SYSTEM FillerModule (* Module Filler, generated from its module specification *)
  (* Standard: 61499-2 *)
  APPLICATION Filler (* Module Filler on target pc (localhost, IO modbus; generated by modgen) *)
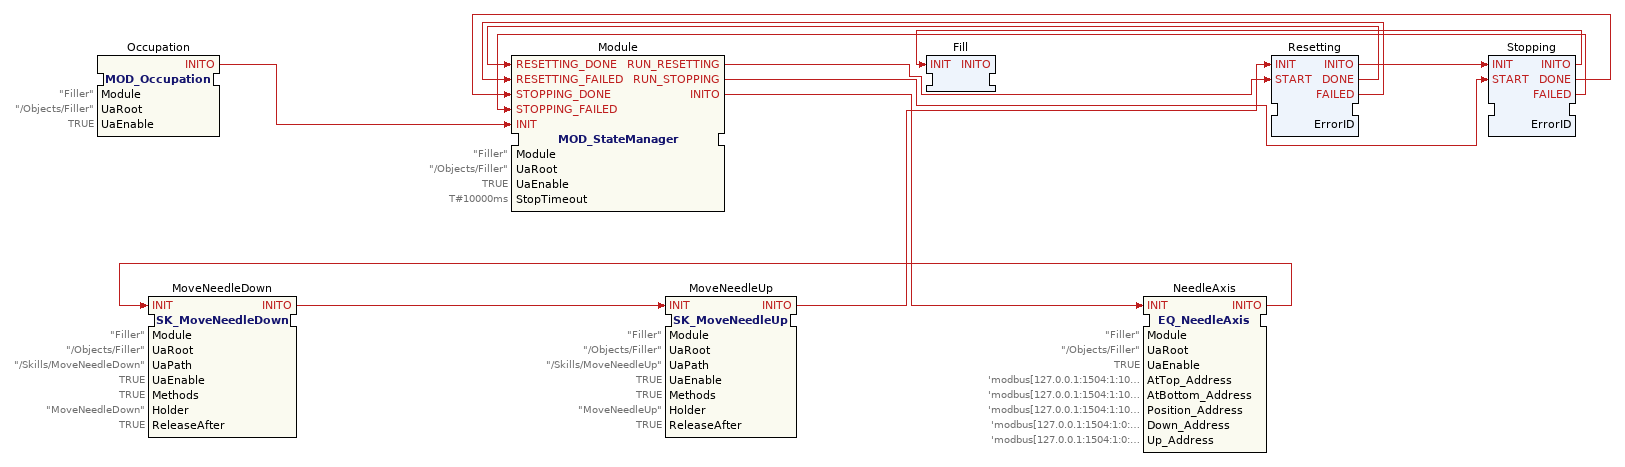
    (* Group ModuleLevel: Module level: occupation, PackML state manager, start-up and the target's IO lines *)
    (* Group ModuleLevelSkills: Module level skills: Control, Sequences (Execute, Stop) of skill primitives and Release; OPC UA /Skills/<name> *)
    (* Group Procedures: Procedures the module state manager runs while Resetting and Stopping *)
    (* Group SkillPrimitives: Skill primitives: one equipment command until a sensor or a time; OPC UA /Skills/<name> *)
    (* Group EquipmentIO: Equipment IO: the only owners of the IO points; skills send them output values over local channels *)
    FBS
      Occupation : modlib::MOD_Occupation(Module := "Filler", UaRoot := "/Objects/Filler", UaEnable := TRUE); (* Who may command the module. A client calls Occupy(Session) at /Objects/Filler/Occupation first; until it calls Release, only commands with that session id are accepted. Every block hears the owner on loc[Filler/owner]. *) {SET_ATTRIBUTE(GroupName, ModuleLevel)}
      Module : modlib::MOD_StateManager(Module := "Filler", UaRoot := "/Objects/Filler", UaEnable := TRUE, StopTimeout := T#10000ms); (* The module's PackML state. The owner calls Reset, Start, Stop, Abort or Clear at /Objects/Filler/Module; State is at /Objects/Filler/Module/State and on loc[Filler/state]. Reset runs the Resetting procedure, Stop the Stopping procedure; skills may be started only in Execute. *) {SET_ATTRIBUTE(GroupName, ModuleLevel)}
      NeedleAxis : filler::EQ_NeedleAxis(Module := "Filler", UaRoot := "/Objects/Filler", UaEnable := TRUE, AtTop_Address := 'modbus[127.0.0.1:1504:1:10:d0:]', AtBottom_Address := 'modbus[127.0.0.1:1504:1:10:d1:]', Position_Address := 'modbus[127.0.0.1:1504:1:10:i1:]', Down_Address := 'modbus[127.0.0.1:1504:1:0::c0]', Up_Address := 'modbus[127.0.0.1:1504:1:0::c2]'); (* Equipment NeedleAxis: Needle lift with down/up valves, end switches and a position sensor. The only block that touches its pins (AtTop = modbus[127.0.0.1:1504:1:10:d0:], AtBottom = modbus[127.0.0.1:1504:1:10:d1:], Position = modbus[127.0.0.1:1504:1:10:i1:], Down = modbus[127.0.0.1:1504:1:0::c0], Up = modbus[127.0.0.1:1504:1:0::c2]). Skills send it what to switch on loc[Filler/NeedleAxis/cmd]; it reports its inputs on loc[Filler/NeedleAxis/state] and at /Objects/Filler/Equipment/NeedleAxis. *) {SET_ATTRIBUTE(GroupName, EquipmentIO)}
      MoveNeedleDown : filler::SK_MoveNeedleDown(Module := "Filler", UaRoot := "/Objects/Filler", UaPath := "/Skills/MoveNeedleDown", UaEnable := TRUE, Methods := TRUE, Holder := "MoveNeedleDown", ReleaseAfter := TRUE); (* Skill MoveNeedleDown, offered on its own: Lower the needle to Distance mm below the top; the default is all the way down, using NeedleAxis. A client calls Start (with the parameters), Stop, Abort or Reset at /Objects/Filler/Skills/MoveNeedleDown; State, ErrorID, Parameters and Results are there too. *) {SET_ATTRIBUTE(GroupName, SkillPrimitives)}
      MoveNeedleUp : filler::SK_MoveNeedleUp(Module := "Filler", UaRoot := "/Objects/Filler", UaPath := "/Skills/MoveNeedleUp", UaEnable := TRUE, Methods := TRUE, Holder := "MoveNeedleUp", ReleaseAfter := TRUE); (* Skill MoveNeedleUp, offered on its own: Raise the needle to the top end switch, using NeedleAxis. A client calls Start (with the parameters), Stop, Abort or Reset at /Objects/Filler/Skills/MoveNeedleUp; State, ErrorID, Parameters and Results are there too. *) {SET_ATTRIBUTE(GroupName, SkillPrimitives)}
    END_FBS
    SUBAPPLICATION Resetting (* Procedure the module runs while Resetting *)
      {SET_ATTRIBUTE(GroupName, Procedures)}
      EVENT_INPUT
        INIT : EInit;
        START;
      END_EVENT
      EVENT_OUTPUT
        INITO : EInit;
        DONE;
        FAILED;
      END_EVENT
      VAR_OUTPUT
        ErrorID : UINT;
      END_VAR
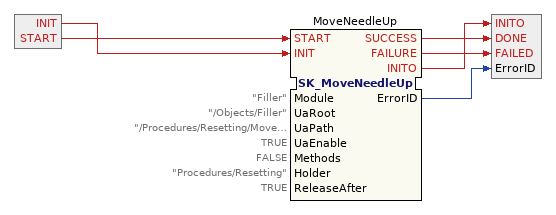
      FBS
        MoveNeedleUp : filler::SK_MoveNeedleUp(Module := "Filler", UaRoot := "/Objects/Filler", UaPath := "/Procedures/Resetting/MoveNeedleUp", UaEnable := TRUE, Methods := FALSE, Holder := "Procedures/Resetting", ReleaseAfter := TRUE); (* Step 1 of Resetting: runs the skill MoveNeedleUp. Its State and ErrorID are at /Objects/Filler/Procedures/Resetting/MoveNeedleUp; it keeps the equipment under the name Procedures/Resetting. *)
      END_FBS
      EVENT_CONNECTIONS
        START TO MoveNeedleUp.START;
        MoveNeedleUp.SUCCESS TO DONE;
        MoveNeedleUp.FAILURE TO FAILED;
        INIT TO MoveNeedleUp.INIT;
        MoveNeedleUp.INITO TO INITO;
      END_CONNECTIONS
      DATA_CONNECTIONS
        MoveNeedleUp.ErrorID TO ErrorID;
      END_CONNECTIONS
    END_SUBAPPLICATION
    SUBAPPLICATION Stopping (* Procedure the module runs while Stopping *)
      {SET_ATTRIBUTE(GroupName, Procedures)}
      EVENT_INPUT
        INIT : EInit;
        START;
      END_EVENT
      EVENT_OUTPUT
        INITO : EInit;
        DONE;
        FAILED;
      END_EVENT
      VAR_OUTPUT
        ErrorID : UINT;
      END_VAR
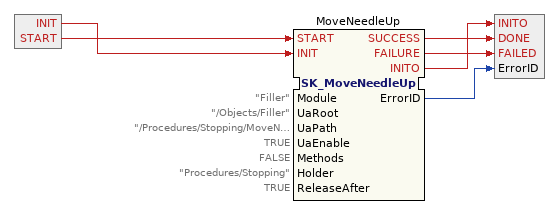
      FBS
        MoveNeedleUp : filler::SK_MoveNeedleUp(Module := "Filler", UaRoot := "/Objects/Filler", UaPath := "/Procedures/Stopping/MoveNeedleUp", UaEnable := TRUE, Methods := FALSE, Holder := "Procedures/Stopping", ReleaseAfter := TRUE); (* Step 1 of Stopping: runs the skill MoveNeedleUp. Its State and ErrorID are at /Objects/Filler/Procedures/Stopping/MoveNeedleUp; it keeps the equipment under the name Procedures/Stopping. *)
      END_FBS
      EVENT_CONNECTIONS
        START TO MoveNeedleUp.START;
        MoveNeedleUp.SUCCESS TO DONE;
        MoveNeedleUp.FAILURE TO FAILED;
        INIT TO MoveNeedleUp.INIT;
        MoveNeedleUp.INITO TO INITO;
      END_CONNECTIONS
      DATA_CONNECTIONS
        MoveNeedleUp.ErrorID TO ErrorID;
      END_CONNECTIONS
    END_SUBAPPLICATION
    SUBAPPLICATION Fill (* Module level skill Fill: Needle down to Depth and back up; a stop lifts the needle *)
      {SET_ATTRIBUTE(GroupName, ModuleLevelSkills)}
      EVENT_INPUT
        INIT : EInit;
      END_EVENT
      EVENT_OUTPUT
        INITO : EInit;
      END_EVENT
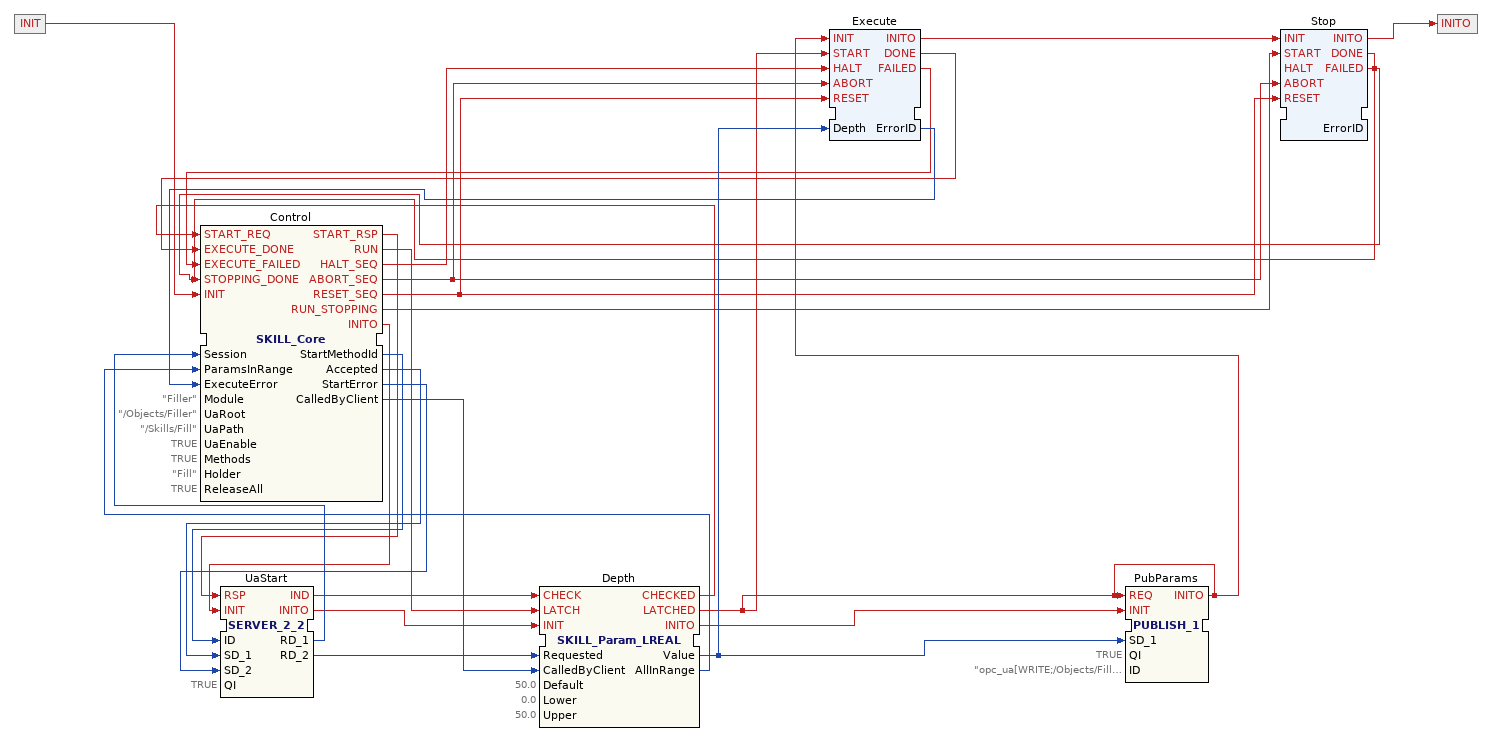
      (* Group Core: The skill's state machine: Stop, Abort, Reset, State and ErrorID over OPC UA; gives up everything the skill holds when a run ends *)
      (* Group Start: The Start method: one block per parameter (range check, value for this run), the values published *)
      (* Group Sequences: What the skill does: Execute, and Stop when it is interrupted; private skill primitives in order *)
      FBS
        Control : modlib::SKILL_Core(Module := "Filler", UaRoot := "/Objects/Filler", UaPath := "/Skills/Fill", UaEnable := TRUE, Methods := TRUE, Holder := "Fill", ReleaseAll := TRUE); (* The state machine of the skill Fill: checks a client's Start (occupation, module in Execute, not running, values in range), publishes State and ErrorID at /Objects/Filler/Skills/Fill, offers Stop, Abort and Reset there, starts Execute and runs Stop when the skill is stopped. *) {SET_ATTRIBUTE(GroupName, Core)}
        UaStart : iec61499::net::SERVER_2_2(QI := TRUE); (* The OPC UA method Start of Fill: a client's call (session id and parameters) arrives here; the parameters are checked, then Control answers Accepted or an error code. *) {SET_ATTRIBUTE(GroupName, Start)}
        Depth : modlib::SKILL_Param_LREAL(Default := 50.0, Lower := 0.0, Upper := 50.0); (* The parameter Depth of Fill: default 50.0 (Lower 0.0, Upper 50.0); checks a client's value, then holds it for the run and hands it to the steps. *) {SET_ATTRIBUTE(GroupName, Start)}
        PubParams : iec61499::net::PUBLISH_1(QI := TRUE, ID := "opc_ua[WRITE;/Objects/Filler/Skills/Fill/Parameters/Depth]"); (* Writes the parameters of the run to OPC UA: /Objects/Filler/Skills/Fill/Parameters/Depth *) {SET_ATTRIBUTE(GroupName, Start)}
      END_FBS
      SUBAPPLICATION Execute (* Fill: execute sequence *)
        {SET_ATTRIBUTE(GroupName, Sequences)}
        EVENT_INPUT
          INIT : EInit;
          START;
          HALT;
          ABORT;
          RESET;
        END_EVENT
        EVENT_OUTPUT
          INITO : EInit;
          DONE;
          FAILED;
        END_EVENT
        VAR_INPUT
          Depth : LREAL;
        END_VAR
        VAR_OUTPUT
          ErrorID : UINT;
        END_VAR
        FBS
          MoveNeedleDown : filler::SK_MoveNeedleDown(Module := "Filler", UaRoot := "/Objects/Filler", UaPath := "/Skills/Fill/Execute/MoveNeedleDown", UaEnable := TRUE, Methods := FALSE, Holder := "Fill", ReleaseAfter := FALSE); (* Step 1 of Fill / Execute: runs the skill MoveNeedleDown; Distance from Fill's Depth. Its State and ErrorID are at /Objects/Filler/Skills/Fill/Execute/MoveNeedleDown; it keeps the equipment under the name Fill. *)
          MoveNeedleUp : filler::SK_MoveNeedleUp(Module := "Filler", UaRoot := "/Objects/Filler", UaPath := "/Skills/Fill/Execute/MoveNeedleUp", UaEnable := TRUE, Methods := FALSE, Holder := "Fill", ReleaseAfter := FALSE); (* Step 2 of Fill / Execute: runs the skill MoveNeedleUp. Its State and ErrorID are at /Objects/Filler/Skills/Fill/Execute/MoveNeedleUp; it keeps the equipment under the name Fill. *)
          Fail1 : modlib::SKILL_FailMerge; (* Joins the failures of the steps into one (with its error code), so any step's failure ends the sequence. *)
        END_FBS
        EVENT_CONNECTIONS
          MoveNeedleDown.SUCCESS TO MoveNeedleUp.START;
          START TO MoveNeedleDown.START;
          MoveNeedleUp.SUCCESS TO DONE;
          MoveNeedleDown.FAILURE TO Fail1.FAIL_1;
          MoveNeedleUp.FAILURE TO Fail1.FAIL_2;
          Fail1.FAIL TO FAILED;
          INIT TO MoveNeedleDown.INIT;
          MoveNeedleUp.INITO TO INITO;
          MoveNeedleDown.INITO TO MoveNeedleUp.INIT;
          HALT TO MoveNeedleDown.HALT;
          HALT TO MoveNeedleUp.HALT;
          ABORT TO MoveNeedleDown.ABORT;
          ABORT TO MoveNeedleUp.ABORT;
          RESET TO MoveNeedleDown.RESET;
          RESET TO MoveNeedleUp.RESET;
        END_CONNECTIONS
        DATA_CONNECTIONS
          Depth TO MoveNeedleDown.Distance;
          MoveNeedleDown.ErrorID TO Fail1.Error1;
          MoveNeedleUp.ErrorID TO Fail1.Error2;
          Fail1.Error TO ErrorID;
        END_CONNECTIONS
      END_SUBAPPLICATION
      SUBAPPLICATION Stop (* Fill: stop sequence *)
        {SET_ATTRIBUTE(GroupName, Sequences)}
        EVENT_INPUT
          INIT : EInit;
          START;
          HALT;
          ABORT;
          RESET;
        END_EVENT
        EVENT_OUTPUT
          INITO : EInit;
          DONE;
          FAILED;
        END_EVENT
        VAR_OUTPUT
          ErrorID : UINT;
        END_VAR
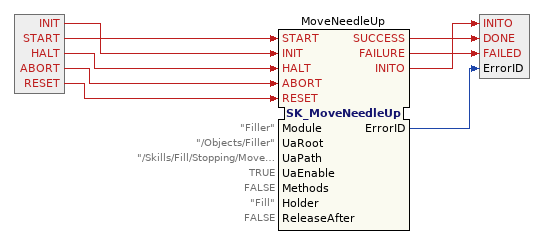
        FBS
          MoveNeedleUp : filler::SK_MoveNeedleUp(Module := "Filler", UaRoot := "/Objects/Filler", UaPath := "/Skills/Fill/Stopping/MoveNeedleUp", UaEnable := TRUE, Methods := FALSE, Holder := "Fill", ReleaseAfter := FALSE); (* Step 1 of Fill / Stop: runs the skill MoveNeedleUp. Its State and ErrorID are at /Objects/Filler/Skills/Fill/Stopping/MoveNeedleUp; it keeps the equipment under the name Fill. *)
        END_FBS
        EVENT_CONNECTIONS
          START TO MoveNeedleUp.START;
          MoveNeedleUp.SUCCESS TO DONE;
          MoveNeedleUp.FAILURE TO FAILED;
          INIT TO MoveNeedleUp.INIT;
          MoveNeedleUp.INITO TO INITO;
          HALT TO MoveNeedleUp.HALT;
          ABORT TO MoveNeedleUp.ABORT;
          RESET TO MoveNeedleUp.RESET;
        END_CONNECTIONS
        DATA_CONNECTIONS
          MoveNeedleUp.ErrorID TO ErrorID;
        END_CONNECTIONS
      END_SUBAPPLICATION
      EVENT_CONNECTIONS
        Control.START_RSP TO UaStart.RSP;
        UaStart.IND TO Depth.CHECK;
        Control.RUN TO Depth.LATCH;
        Depth.CHECKED TO Control.START_REQ;
        Depth.LATCHED TO PubParams.REQ;
        PubParams.INITO TO PubParams.REQ;
        Depth.LATCHED TO Execute.START;
        Control.HALT_SEQ TO Execute.HALT;
        Control.ABORT_SEQ TO Execute.ABORT;
        Control.RESET_SEQ TO Execute.RESET;
        Execute.DONE TO Control.EXECUTE_DONE;
        Execute.FAILED TO Control.EXECUTE_FAILED;
        Control.RUN_STOPPING TO Stop.START;
        Control.ABORT_SEQ TO Stop.ABORT;
        Control.RESET_SEQ TO Stop.RESET;
        Stop.DONE TO Control.STOPPING_DONE;
        Stop.FAILED TO Control.STOPPING_DONE;
        INIT TO Control.INIT;
        Control.INITO TO UaStart.INIT;
        UaStart.INITO TO Depth.INIT;
        Depth.INITO TO PubParams.INIT;
        PubParams.INITO TO Execute.INIT;
        Execute.INITO TO Stop.INIT;
        Stop.INITO TO INITO;
      END_CONNECTIONS
      DATA_CONNECTIONS
        Control.StartMethodId TO UaStart.ID;
        UaStart.RD_1 TO Control.Session;
        Control.Accepted TO UaStart.SD_1;
        Control.StartError TO UaStart.SD_2;
        UaStart.RD_2 TO Depth.Requested;
        Control.CalledByClient TO Depth.CalledByClient;
        Depth.Value TO PubParams.SD_1;
        Depth.AllInRange TO Control.ParamsInRange;
        Depth.Value TO Execute.Depth;
        Execute.ErrorID TO Control.ExecuteError;
      END_CONNECTIONS
    END_SUBAPPLICATION
    EVENT_CONNECTIONS
      Module.RUN_RESETTING TO Resetting.START;
      Resetting.DONE TO Module.RESETTING_DONE;
      Resetting.FAILED TO Module.RESETTING_FAILED;
      Module.RUN_STOPPING TO Stopping.START;
      Stopping.DONE TO Module.STOPPING_DONE;
      Stopping.FAILED TO Module.STOPPING_FAILED;
      Occupation.INITO TO Module.INIT;
      Module.INITO TO NeedleAxis.INIT;
      NeedleAxis.INITO TO MoveNeedleDown.INIT;
      MoveNeedleDown.INITO TO MoveNeedleUp.INIT;
      MoveNeedleUp.INITO TO Resetting.INIT;
      Resetting.INITO TO Stopping.INIT;
      Stopping.INITO TO Fill.INIT;
    END_CONNECTIONS
  END_APPLICATION
  APPLICATION Filler_pi (* Module Filler on target pi (filler-pi.invalid, IO gpio; generated by modgen) *)
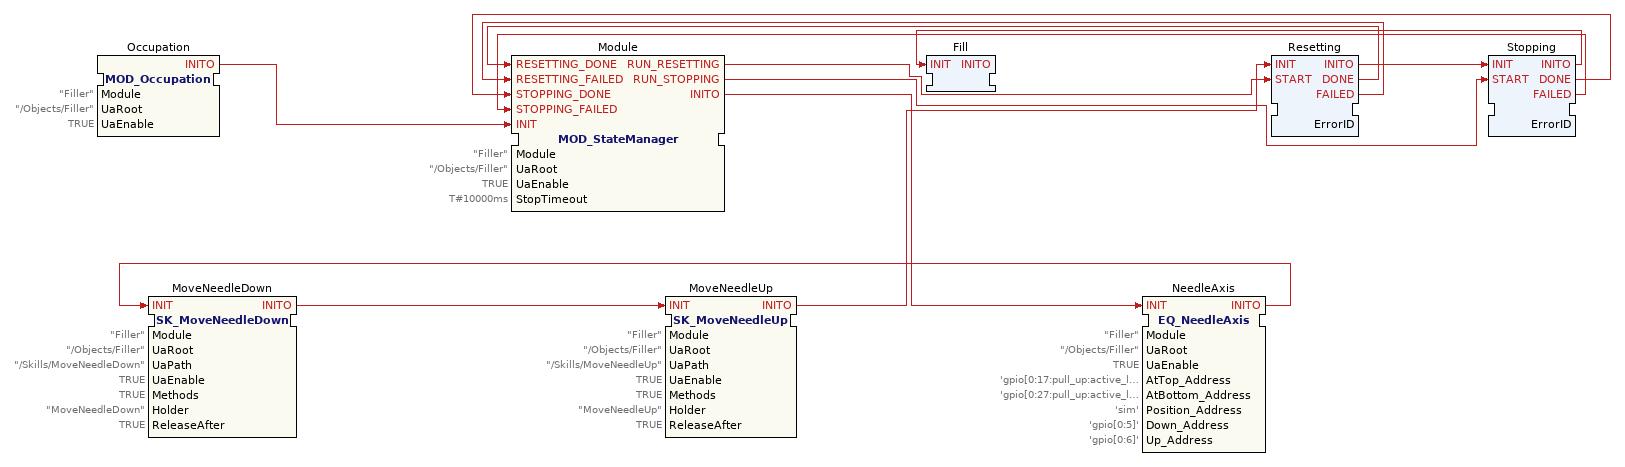
    (* Group ModuleLevel: Module level: occupation, PackML state manager, start-up and the target's IO lines *)
    (* Group ModuleLevelSkills: Module level skills: Control, Sequences (Execute, Stop) of skill primitives and Release; OPC UA /Skills/<name> *)
    (* Group Procedures: Procedures the module state manager runs while Resetting and Stopping *)
    (* Group SkillPrimitives: Skill primitives: one equipment command until a sensor or a time; OPC UA /Skills/<name> *)
    (* Group EquipmentIO: Equipment IO: the only owners of the IO points; skills send them output values over local channels *)
    FBS
      Occupation : modlib::MOD_Occupation(Module := "Filler", UaRoot := "/Objects/Filler", UaEnable := TRUE); (* Who may command the module. A client calls Occupy(Session) at /Objects/Filler/Occupation first; until it calls Release, only commands with that session id are accepted. Every block hears the owner on loc[Filler/owner]. *) {SET_ATTRIBUTE(GroupName, ModuleLevel)}
      Module : modlib::MOD_StateManager(Module := "Filler", UaRoot := "/Objects/Filler", UaEnable := TRUE, StopTimeout := T#10000ms); (* The module's PackML state. The owner calls Reset, Start, Stop, Abort or Clear at /Objects/Filler/Module; State is at /Objects/Filler/Module/State and on loc[Filler/state]. Reset runs the Resetting procedure, Stop the Stopping procedure; skills may be started only in Execute. *) {SET_ATTRIBUTE(GroupName, ModuleLevel)}
      NeedleAxis : filler::EQ_NeedleAxis(Module := "Filler", UaRoot := "/Objects/Filler", UaEnable := TRUE, AtTop_Address := 'gpio[0:17:pull_up:active_low]', AtBottom_Address := 'gpio[0:27:pull_up:active_low]', Position_Address := 'sim', Down_Address := 'gpio[0:5]', Up_Address := 'gpio[0:6]'); (* Equipment NeedleAxis: Needle lift with down/up valves, end switches and a position sensor. The only block that touches its pins (AtTop = gpio[0:17:pull_up:active_low], AtBottom = gpio[0:27:pull_up:active_low], Position = sim, Down = gpio[0:5], Up = gpio[0:6]). Skills send it what to switch on loc[Filler/NeedleAxis/cmd]; it reports its inputs on loc[Filler/NeedleAxis/state] and at /Objects/Filler/Equipment/NeedleAxis. *) {SET_ATTRIBUTE(GroupName, EquipmentIO)}
      MoveNeedleDown : filler::SK_MoveNeedleDown(Module := "Filler", UaRoot := "/Objects/Filler", UaPath := "/Skills/MoveNeedleDown", UaEnable := TRUE, Methods := TRUE, Holder := "MoveNeedleDown", ReleaseAfter := TRUE); (* Skill MoveNeedleDown, offered on its own: Lower the needle to Distance mm below the top; the default is all the way down, using NeedleAxis. A client calls Start (with the parameters), Stop, Abort or Reset at /Objects/Filler/Skills/MoveNeedleDown; State, ErrorID, Parameters and Results are there too. *) {SET_ATTRIBUTE(GroupName, SkillPrimitives)}
      MoveNeedleUp : filler::SK_MoveNeedleUp(Module := "Filler", UaRoot := "/Objects/Filler", UaPath := "/Skills/MoveNeedleUp", UaEnable := TRUE, Methods := TRUE, Holder := "MoveNeedleUp", ReleaseAfter := TRUE); (* Skill MoveNeedleUp, offered on its own: Raise the needle to the top end switch, using NeedleAxis. A client calls Start (with the parameters), Stop, Abort or Reset at /Objects/Filler/Skills/MoveNeedleUp; State, ErrorID, Parameters and Results are there too. *) {SET_ATTRIBUTE(GroupName, SkillPrimitives)}
    END_FBS
    SUBAPPLICATION Resetting (* Procedure the module runs while Resetting *)
      {SET_ATTRIBUTE(GroupName, Procedures)}
      EVENT_INPUT
        INIT : EInit;
        START;
      END_EVENT
      EVENT_OUTPUT
        INITO : EInit;
        DONE;
        FAILED;
      END_EVENT
      VAR_OUTPUT
        ErrorID : UINT;
      END_VAR
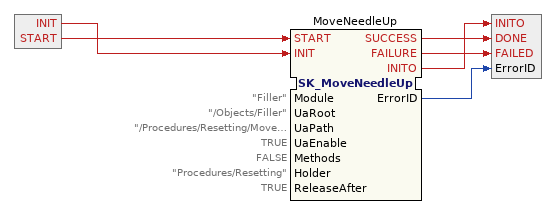
      FBS
        MoveNeedleUp : filler::SK_MoveNeedleUp(Module := "Filler", UaRoot := "/Objects/Filler", UaPath := "/Procedures/Resetting/MoveNeedleUp", UaEnable := TRUE, Methods := FALSE, Holder := "Procedures/Resetting", ReleaseAfter := TRUE); (* Step 1 of Resetting: runs the skill MoveNeedleUp. Its State and ErrorID are at /Objects/Filler/Procedures/Resetting/MoveNeedleUp; it keeps the equipment under the name Procedures/Resetting. *)
      END_FBS
      EVENT_CONNECTIONS
        START TO MoveNeedleUp.START;
        MoveNeedleUp.SUCCESS TO DONE;
        MoveNeedleUp.FAILURE TO FAILED;
        INIT TO MoveNeedleUp.INIT;
        MoveNeedleUp.INITO TO INITO;
      END_CONNECTIONS
      DATA_CONNECTIONS
        MoveNeedleUp.ErrorID TO ErrorID;
      END_CONNECTIONS
    END_SUBAPPLICATION
    SUBAPPLICATION Stopping (* Procedure the module runs while Stopping *)
      {SET_ATTRIBUTE(GroupName, Procedures)}
      EVENT_INPUT
        INIT : EInit;
        START;
      END_EVENT
      EVENT_OUTPUT
        INITO : EInit;
        DONE;
        FAILED;
      END_EVENT
      VAR_OUTPUT
        ErrorID : UINT;
      END_VAR
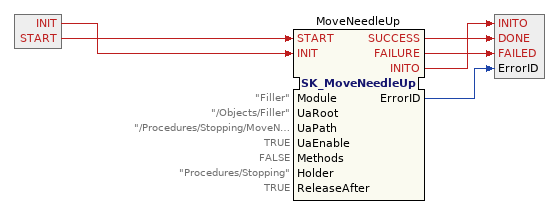
      FBS
        MoveNeedleUp : filler::SK_MoveNeedleUp(Module := "Filler", UaRoot := "/Objects/Filler", UaPath := "/Procedures/Stopping/MoveNeedleUp", UaEnable := TRUE, Methods := FALSE, Holder := "Procedures/Stopping", ReleaseAfter := TRUE); (* Step 1 of Stopping: runs the skill MoveNeedleUp. Its State and ErrorID are at /Objects/Filler/Procedures/Stopping/MoveNeedleUp; it keeps the equipment under the name Procedures/Stopping. *)
      END_FBS
      EVENT_CONNECTIONS
        START TO MoveNeedleUp.START;
        MoveNeedleUp.SUCCESS TO DONE;
        MoveNeedleUp.FAILURE TO FAILED;
        INIT TO MoveNeedleUp.INIT;
        MoveNeedleUp.INITO TO INITO;
      END_CONNECTIONS
      DATA_CONNECTIONS
        MoveNeedleUp.ErrorID TO ErrorID;
      END_CONNECTIONS
    END_SUBAPPLICATION
    SUBAPPLICATION Fill (* Module level skill Fill: Needle down to Depth and back up; a stop lifts the needle *)
      {SET_ATTRIBUTE(GroupName, ModuleLevelSkills)}
      EVENT_INPUT
        INIT : EInit;
      END_EVENT
      EVENT_OUTPUT
        INITO : EInit;
      END_EVENT
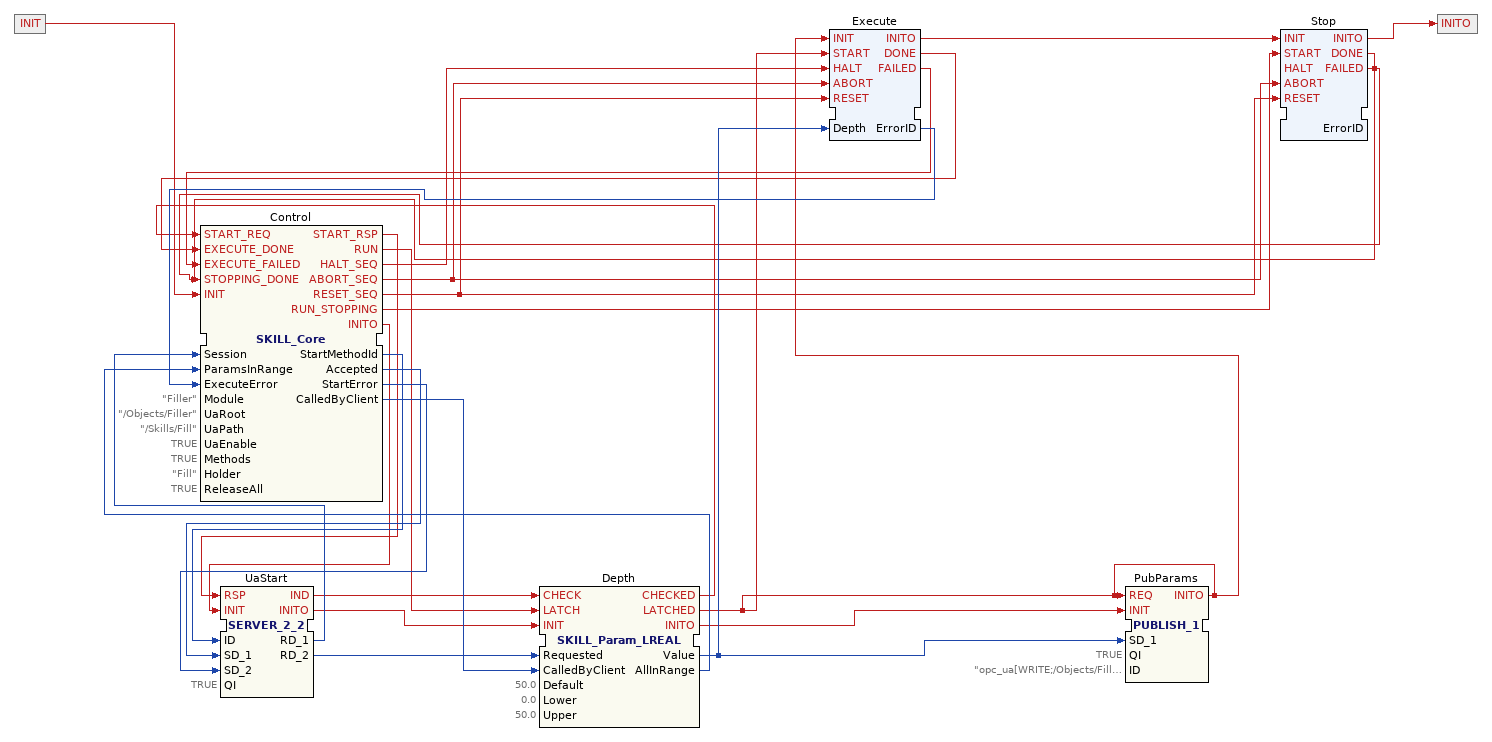
      (* Group Core: The skill's state machine: Stop, Abort, Reset, State and ErrorID over OPC UA; gives up everything the skill holds when a run ends *)
      (* Group Start: The Start method: one block per parameter (range check, value for this run), the values published *)
      (* Group Sequences: What the skill does: Execute, and Stop when it is interrupted; private skill primitives in order *)
      FBS
        Control : modlib::SKILL_Core(Module := "Filler", UaRoot := "/Objects/Filler", UaPath := "/Skills/Fill", UaEnable := TRUE, Methods := TRUE, Holder := "Fill", ReleaseAll := TRUE); (* The state machine of the skill Fill: checks a client's Start (occupation, module in Execute, not running, values in range), publishes State and ErrorID at /Objects/Filler/Skills/Fill, offers Stop, Abort and Reset there, starts Execute and runs Stop when the skill is stopped. *) {SET_ATTRIBUTE(GroupName, Core)}
        UaStart : iec61499::net::SERVER_2_2(QI := TRUE); (* The OPC UA method Start of Fill: a client's call (session id and parameters) arrives here; the parameters are checked, then Control answers Accepted or an error code. *) {SET_ATTRIBUTE(GroupName, Start)}
        Depth : modlib::SKILL_Param_LREAL(Default := 50.0, Lower := 0.0, Upper := 50.0); (* The parameter Depth of Fill: default 50.0 (Lower 0.0, Upper 50.0); checks a client's value, then holds it for the run and hands it to the steps. *) {SET_ATTRIBUTE(GroupName, Start)}
        PubParams : iec61499::net::PUBLISH_1(QI := TRUE, ID := "opc_ua[WRITE;/Objects/Filler/Skills/Fill/Parameters/Depth]"); (* Writes the parameters of the run to OPC UA: /Objects/Filler/Skills/Fill/Parameters/Depth *) {SET_ATTRIBUTE(GroupName, Start)}
      END_FBS
      SUBAPPLICATION Execute (* Fill: execute sequence *)
        {SET_ATTRIBUTE(GroupName, Sequences)}
        EVENT_INPUT
          INIT : EInit;
          START;
          HALT;
          ABORT;
          RESET;
        END_EVENT
        EVENT_OUTPUT
          INITO : EInit;
          DONE;
          FAILED;
        END_EVENT
        VAR_INPUT
          Depth : LREAL;
        END_VAR
        VAR_OUTPUT
          ErrorID : UINT;
        END_VAR
        FBS
          MoveNeedleDown : filler::SK_MoveNeedleDown(Module := "Filler", UaRoot := "/Objects/Filler", UaPath := "/Skills/Fill/Execute/MoveNeedleDown", UaEnable := TRUE, Methods := FALSE, Holder := "Fill", ReleaseAfter := FALSE); (* Step 1 of Fill / Execute: runs the skill MoveNeedleDown; Distance from Fill's Depth. Its State and ErrorID are at /Objects/Filler/Skills/Fill/Execute/MoveNeedleDown; it keeps the equipment under the name Fill. *)
          MoveNeedleUp : filler::SK_MoveNeedleUp(Module := "Filler", UaRoot := "/Objects/Filler", UaPath := "/Skills/Fill/Execute/MoveNeedleUp", UaEnable := TRUE, Methods := FALSE, Holder := "Fill", ReleaseAfter := FALSE); (* Step 2 of Fill / Execute: runs the skill MoveNeedleUp. Its State and ErrorID are at /Objects/Filler/Skills/Fill/Execute/MoveNeedleUp; it keeps the equipment under the name Fill. *)
          Fail1 : modlib::SKILL_FailMerge; (* Joins the failures of the steps into one (with its error code), so any step's failure ends the sequence. *)
        END_FBS
        EVENT_CONNECTIONS
          MoveNeedleDown.SUCCESS TO MoveNeedleUp.START;
          START TO MoveNeedleDown.START;
          MoveNeedleUp.SUCCESS TO DONE;
          MoveNeedleDown.FAILURE TO Fail1.FAIL_1;
          MoveNeedleUp.FAILURE TO Fail1.FAIL_2;
          Fail1.FAIL TO FAILED;
          INIT TO MoveNeedleDown.INIT;
          MoveNeedleUp.INITO TO INITO;
          MoveNeedleDown.INITO TO MoveNeedleUp.INIT;
          HALT TO MoveNeedleDown.HALT;
          HALT TO MoveNeedleUp.HALT;
          ABORT TO MoveNeedleDown.ABORT;
          ABORT TO MoveNeedleUp.ABORT;
          RESET TO MoveNeedleDown.RESET;
          RESET TO MoveNeedleUp.RESET;
        END_CONNECTIONS
        DATA_CONNECTIONS
          Depth TO MoveNeedleDown.Distance;
          MoveNeedleDown.ErrorID TO Fail1.Error1;
          MoveNeedleUp.ErrorID TO Fail1.Error2;
          Fail1.Error TO ErrorID;
        END_CONNECTIONS
      END_SUBAPPLICATION
      SUBAPPLICATION Stop (* Fill: stop sequence *)
        {SET_ATTRIBUTE(GroupName, Sequences)}
        EVENT_INPUT
          INIT : EInit;
          START;
          HALT;
          ABORT;
          RESET;
        END_EVENT
        EVENT_OUTPUT
          INITO : EInit;
          DONE;
          FAILED;
        END_EVENT
        VAR_OUTPUT
          ErrorID : UINT;
        END_VAR
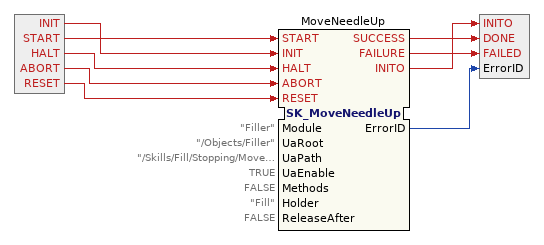
        FBS
          MoveNeedleUp : filler::SK_MoveNeedleUp(Module := "Filler", UaRoot := "/Objects/Filler", UaPath := "/Skills/Fill/Stopping/MoveNeedleUp", UaEnable := TRUE, Methods := FALSE, Holder := "Fill", ReleaseAfter := FALSE); (* Step 1 of Fill / Stop: runs the skill MoveNeedleUp. Its State and ErrorID are at /Objects/Filler/Skills/Fill/Stopping/MoveNeedleUp; it keeps the equipment under the name Fill. *)
        END_FBS
        EVENT_CONNECTIONS
          START TO MoveNeedleUp.START;
          MoveNeedleUp.SUCCESS TO DONE;
          MoveNeedleUp.FAILURE TO FAILED;
          INIT TO MoveNeedleUp.INIT;
          MoveNeedleUp.INITO TO INITO;
          HALT TO MoveNeedleUp.HALT;
          ABORT TO MoveNeedleUp.ABORT;
          RESET TO MoveNeedleUp.RESET;
        END_CONNECTIONS
        DATA_CONNECTIONS
          MoveNeedleUp.ErrorID TO ErrorID;
        END_CONNECTIONS
      END_SUBAPPLICATION
      EVENT_CONNECTIONS
        Control.START_RSP TO UaStart.RSP;
        UaStart.IND TO Depth.CHECK;
        Control.RUN TO Depth.LATCH;
        Depth.CHECKED TO Control.START_REQ;
        Depth.LATCHED TO PubParams.REQ;
        PubParams.INITO TO PubParams.REQ;
        Depth.LATCHED TO Execute.START;
        Control.HALT_SEQ TO Execute.HALT;
        Control.ABORT_SEQ TO Execute.ABORT;
        Control.RESET_SEQ TO Execute.RESET;
        Execute.DONE TO Control.EXECUTE_DONE;
        Execute.FAILED TO Control.EXECUTE_FAILED;
        Control.RUN_STOPPING TO Stop.START;
        Control.ABORT_SEQ TO Stop.ABORT;
        Control.RESET_SEQ TO Stop.RESET;
        Stop.DONE TO Control.STOPPING_DONE;
        Stop.FAILED TO Control.STOPPING_DONE;
        INIT TO Control.INIT;
        Control.INITO TO UaStart.INIT;
        UaStart.INITO TO Depth.INIT;
        Depth.INITO TO PubParams.INIT;
        PubParams.INITO TO Execute.INIT;
        Execute.INITO TO Stop.INIT;
        Stop.INITO TO INITO;
      END_CONNECTIONS
      DATA_CONNECTIONS
        Control.StartMethodId TO UaStart.ID;
        UaStart.RD_1 TO Control.Session;
        Control.Accepted TO UaStart.SD_1;
        Control.StartError TO UaStart.SD_2;
        UaStart.RD_2 TO Depth.Requested;
        Control.CalledByClient TO Depth.CalledByClient;
        Depth.Value TO PubParams.SD_1;
        Depth.AllInRange TO Control.ParamsInRange;
        Depth.Value TO Execute.Depth;
        Execute.ErrorID TO Control.ExecuteError;
      END_CONNECTIONS
    END_SUBAPPLICATION
    EVENT_CONNECTIONS
      Module.RUN_RESETTING TO Resetting.START;
      Resetting.DONE TO Module.RESETTING_DONE;
      Resetting.FAILED TO Module.RESETTING_FAILED;
      Module.RUN_STOPPING TO Stopping.START;
      Stopping.DONE TO Module.STOPPING_DONE;
      Stopping.FAILED TO Module.STOPPING_FAILED;
      Occupation.INITO TO Module.INIT;
      Module.INITO TO NeedleAxis.INIT;
      NeedleAxis.INITO TO MoveNeedleDown.INIT;
      MoveNeedleDown.INITO TO MoveNeedleUp.INIT;
      MoveNeedleUp.INITO TO Resetting.INIT;
      Resetting.INITO TO Stopping.INIT;
      Stopping.INITO TO Fill.INIT;
    END_CONNECTIONS
  END_APPLICATION
  DEVICE FORTE_PC : iec61499::system::FORTE_PC(MGR_ID := "localhost:61499" (* Device manager socket ID *))
    {SET_ATTRIBUTE(Profile, HOLOBLOC)}
    RESOURCE RES : iec61499::system::EMB_RES
      EVENT_CONNECTIONS
        START.COLD TO Filler.Occupation.INIT;
        START.WARM TO Filler.Occupation.INIT;
      END_CONNECTIONS
    END_RESOURCE
  END_DEVICE
  DEVICE FORTE_PI : iec61499::system::FORTE_PC(MGR_ID := "filler-pi.invalid:61499" (* Device manager socket ID *))
    {SET_ATTRIBUTE(Profile, HOLOBLOC)}
    RESOURCE RES : iec61499::system::EMB_RES
      EVENT_CONNECTIONS
        START.COLD TO Filler_pi.Occupation.INIT;
        START.WARM TO Filler_pi.Occupation.INIT;
      END_CONNECTIONS
    END_RESOURCE
  END_DEVICE
  MAPPINGS
    Filler.Occupation ON FORTE_PC.RES;
    Filler.Module ON FORTE_PC.RES;
    Filler.NeedleAxis ON FORTE_PC.RES;
    Filler.MoveNeedleDown ON FORTE_PC.RES;
    Filler.MoveNeedleUp ON FORTE_PC.RES;
    Filler.Resetting ON FORTE_PC.RES;
    Filler.Stopping ON FORTE_PC.RES;
    Filler.Fill ON FORTE_PC.RES;
    Filler_pi.Occupation ON FORTE_PI.RES;
    Filler_pi.Module ON FORTE_PI.RES;
    Filler_pi.NeedleAxis ON FORTE_PI.RES;
    Filler_pi.MoveNeedleDown ON FORTE_PI.RES;
    Filler_pi.MoveNeedleUp ON FORTE_PI.RES;
    Filler_pi.Resetting ON FORTE_PI.RES;
    Filler_pi.Stopping ON FORTE_PI.RES;
    Filler_pi.Fill ON FORTE_PI.RES;
  END_MAPPINGS
END_SYSTEM
